// Generated by voz_llm_plc_agent
// Target: Siemens TIA Portal V18 - SCL external source
// Review and compile before any download to physical hardware.

FUNCTION_BLOCK "PLC_PRG"
{ S7_Optimized_Access := 'TRUE' }
VERSION : 0.1
VAR_INPUT
   I_Speed_Low : Bool := FALSE;
   I_Speed_Medium : Bool := FALSE;
   I_Speed_High : Bool := FALSE;
   I_Emergency : Bool := FALSE;
END_VAR
VAR_OUTPUT
   Q_Speed_Low : Bool := FALSE;
   Q_Speed_Medium : Bool := FALSE;
   Q_Speed_High : Bool := FALSE;
END_VAR
BEGIN
(* Seleccion de velocidad: solo se activa la velocidad seleccionada; con mas de una seleccion *)
(* simultanea ninguna se activa (nunca dos velocidades a la vez). *)
#Q_Speed_Low := #I_Speed_Low AND NOT #I_Speed_Medium AND NOT #I_Speed_High AND NOT #I_Emergency;
#Q_Speed_Medium := #I_Speed_Medium AND NOT #I_Speed_Low AND NOT #I_Speed_High AND NOT #I_Emergency;
#Q_Speed_High := #I_Speed_High AND NOT #I_Speed_Low AND NOT #I_Speed_Medium AND NOT #I_Emergency;
END_FUNCTION_BLOCK

DATA_BLOCK "DB_PLC_PRG"
{ S7_Optimized_Access := 'TRUE' }
VERSION : 0.1
NON_RETAIN
"PLC_PRG"
BEGIN
END_DATA_BLOCK

ORGANIZATION_BLOCK "Main"
{ S7_Optimized_Access := 'TRUE' }
VERSION : 0.1
BEGIN
   "DB_PLC_PRG"(
      I_Speed_Low := "I_Speed_Low",
      I_Speed_Medium := "I_Speed_Medium",
      I_Speed_High := "I_Speed_High",
      I_Emergency := "I_Emergency",
      Q_Speed_Low => "Q_Speed_Low",
      Q_Speed_Medium => "Q_Speed_Medium",
      Q_Speed_High => "Q_Speed_High"
   );
END_ORGANIZATION_BLOCK
